(* IEC 61131-3 sources: CannyIECUnitTest/st/device/plc_logic/application, 5 files *)

(* ---- testcase-TestCase.st ---- *)
(* --- Interface --- *)
{attribute 'test'}
{attribute 'testcasetimeout':='15000'}
FUNCTION_BLOCK TestCase EXTENDS TM.Testcase
VAR_INPUT
END_VAR
VAR_OUTPUT
END_VAR
VAR
END_VAR

(* --- Implementation --- *)
SUPER^();

(* ---- testcase_consheap-TestCase_ConsHeap.st ---- *)
(* --- Interface --- *)
{attribute 'test'}
{attribute 'testcasename':='ConsHeap'}
{attribute 'testcasetimeout':='15000'}
FUNCTION_BLOCK TestCase_ConsHeap EXTENDS Testcase
VAR_INPUT
END_VAR
VAR_OUTPUT
END_VAR
VAR
END_VAR

(* --- Implementation --- *)
SUPER^();

(* ---- testcase_isignbit-TestCase_ISIGNBIT.st ---- *)
(* --- Interface --- *)
{attribute 'test'}
{attribute 'testcasename':='ISIGNBIT'}
{attribute 'testcasetimeout':='15000'}
FUNCTION_BLOCK TestCase_ISIGNBIT EXTENDS Testcase
VAR_INPUT
END_VAR
VAR_OUTPUT
END_VAR
VAR
END_VAR

(* --- Implementation --- *)
SUPER^();

(* ---- testcase_loadbank-TestCase_LoadBank.st ---- *)
(* --- Interface --- *)
{attribute 'test'}
{attribute 'testcasename':='LoadBank'}
{attribute 'testcasetimeout':='15000'}
FUNCTION_BLOCK TestCase_LoadBank EXTENDS Testcase
VAR_INPUT
END_VAR
VAR_OUTPUT
END_VAR
VAR
END_VAR

(* --- Implementation --- *)
SUPER^();

(* ---- plc_prg-PLC_PRG.st ---- *)
(* --- Interface --- *)
PROGRAM PLC_PRG
VAR
	fbTestCase_ISIGNBIT : TestCase_ISIGNBIT;
	fbTestCase_ConsHeap : TestCase_ConsHeap;
	fbTestCase_LoadBank : TestCase_LoadBank;
END_VAR
